Fanuc KAREL source: KA00213.KL

PROGRAM KA00213
%NOLOCKGROUP
VAR
  SRC: ARRAY[4] OF XYZWPR
  DST: ARRAY[4] OF SHORT
BEGIN
  DST = SRC
END KA00213
